{attribute 'pack_mode' := '1'}
TYPE ST_TRIGERS_StrengthAnalysis :
STRUCT
	
	sHMI_Mode									: STRING(254);
	bControlOn									: BOOL;	//kluczyk-sterowanie załączone
	bCycleStartCmd								: BOOL;	//przycisk start cyklu
	bCycleStopCmd								: BOOL;	//przycisk stop cyklu
	bAutoMode									: BOOL;	//tryb automatyczny
	bBreakthroughDetection_2_BreakDetected		: BOOL;
	//arrEHS_EventVisu							: ARRAY [1..GVL_EHS.diNoOfEvents] OF ST_EventHistoricalSimple;	

END_STRUCT
END_TYPE

(* stored: Version 1.1.0.1, ProductVersion 3.1.4024.15
   DUT ST_TRIGERS_StrengthAnalysis: Id {058aaf0f-f5e3-423e-9386-6938de1b98ad} *)
